(* IEC 61131-3 sources: codesys-api/examples/codesys4/projects/modbus_probe.fbsdev/Application.iecapp^, 1 file *)

(* ---- PLC_PRG.prg.st ---- *)
PROGRAM PLC_PRG
VAR
    counter : INT;
    flag : BOOL;
END_VAR
counter := counter + 1;
flag := counter > 10;
END_PROGRAM
